Fanuc KAREL source: KA00008.KL

PROGRAM KA00008
%NOLOCKGROUP
VAR
  SRC: INTEGER
  DST: JOINTPOS
BEGIN
  SRC = 2
  DST = SRC
END KA00008
